Fanuc KAREL source: KT00514.KL

PROGRAM KT00514
%NOLOCKGROUP
VAR
  P1: XYZWPREXT
  P2: POSITION
  OUT: POSITION
BEGIN
  P1.X = 1.0
  OUT = P1 : P2
END KT00514
